FUNCTION_BLOCK FB_DriveStatus (* Migrated from IEC 61131-3 ST *)
  (* Standard: 61499-2 *)
  (* Version 1.0, 2026-11-06, st2fb *)
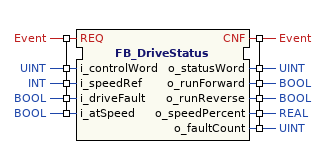
  EVENT_INPUT
    REQ WITH i_controlWord, i_speedRef, i_driveFault, i_atSpeed;
  END_EVENT
  EVENT_OUTPUT
    CNF WITH o_statusWord, o_runForward, o_runReverse, o_speedPercent, o_faultCount;
  END_EVENT
  VAR_INPUT
    i_controlWord : UINT;
    i_speedRef : INT;
    i_driveFault : BOOL;
    i_atSpeed : BOOL;
  END_VAR
  VAR_OUTPUT
    o_statusWord : UINT;
    o_runForward : BOOL;
    o_runReverse : BOOL;
    o_speedPercent : REAL;
    o_faultCount : UINT;
  END_VAR
  VAR
    statFaultLatched : BOOL := FALSE;
    statFaultEdge_CLK : BOOL := FALSE;
    statFaultEdge_Q : BOOL := FALSE;
    statFaultEdge_M : BOOL := FALSE;
  END_VAR
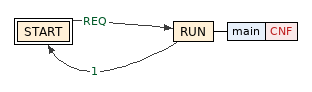
  EC_STATES
    START;
    RUN : main -> CNF;
  END_STATES
  EC_TRANSITIONS
    START TO RUN := REQ;
    RUN TO START := 1;
  END_TRANSITIONS
  ALGORITHM main IN ST:
statFaultEdge_CLK := i_driveFault;
statFaultEdge_Q := statFaultEdge_CLK AND NOT statFaultEdge_M;
statFaultEdge_M := statFaultEdge_CLK;
IF statFaultEdge_Q THEN
  o_faultCount := o_faultCount + 1;
END_IF;
IF i_driveFault THEN
  statFaultLatched := TRUE;
ELSIF (UINT_TO_INT(i_controlWord / 128) MOD 2) = 1 THEN
  statFaultLatched := FALSE;
END_IF;
o_runForward := ((i_controlWord MOD 2) = 1) AND ((UINT_TO_INT(i_controlWord / 2) MOD 2) = 1) AND NOT ((UINT_TO_INT(i_controlWord / 4) MOD 2) = 1) AND NOT statFaultLatched;
o_runReverse := ((i_controlWord MOD 2) = 1) AND ((UINT_TO_INT(i_controlWord / 2) MOD 2) = 1) AND ((UINT_TO_INT(i_controlWord / 4) MOD 2) = 1) AND NOT statFaultLatched;
IF o_runForward OR o_runReverse THEN
  o_speedPercent := INT_TO_REAL(i_speedRef) * 100.0 / 16384.0;
ELSE
  o_speedPercent := 0.0;
END_IF;
o_statusWord := 0;
IF ((i_controlWord MOD 2) = 1) AND NOT statFaultLatched THEN
  o_statusWord := o_statusWord + 1;
END_IF;
IF o_runForward OR o_runReverse THEN
  o_statusWord := o_statusWord + 2;
END_IF;
IF o_runReverse THEN
  o_statusWord := o_statusWord + 4;
END_IF;
IF statFaultLatched THEN
  o_statusWord := o_statusWord + 8;
END_IF;
IF i_atSpeed AND (o_runForward OR o_runReverse) THEN
  o_statusWord := o_statusWord + 16;
END_IF;
  END_ALGORITHM
END_FUNCTION_BLOCK
